// LS Electric XG5000 project: COMFactoryIO_Automated Warehouse10TL
// PLC LSPLC

PROGRAM NewProgram (task: 스캔 프로그램)

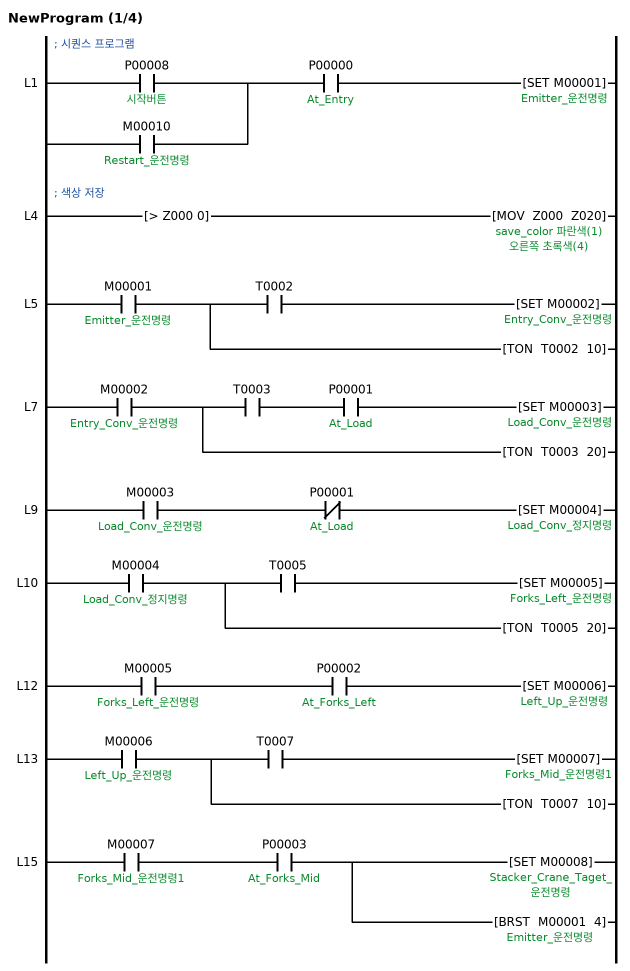
// 시퀀스 프로그램
; L1
LOAD      P00008	// 시작버튼
OR        M00010	// Restart_운전명령
AND       P00000	// At_Entry
SET       M00001	// Emitter_운전명령
// 색상 저장
; L4
LOAD>     Z000 0
MOV       Z000 Z020	// save_color 파란색(1) 오른쪽 초록색(4)
; L5
LOAD      M00001	// Emitter_운전명령
MPUSH
AND       T0002
SET       M00002	// Entry_Conv_운전명령
MPOP
TON       T0002 10
; L7
LOAD      M00002	// Entry_Conv_운전명령
MPUSH
AND       T0003
AND       P00001	// At_Load
SET       M00003	// Load_Conv_운전명령
MPOP
TON       T0003 20
; L9
LOAD      M00003	// Load_Conv_운전명령
AND NOT   P00001	// At_Load
SET       M00004	// Load_Conv_정지명령
; L10
LOAD      M00004	// Load_Conv_정지명령
MPUSH
AND       T0005
SET       M00005	// Forks_Left_운전명령
MPOP
TON       T0005 20
; L12
LOAD      M00005	// Forks_Left_운전명령
AND       P00002	// At_Forks_Left
SET       M00006	// Left_Up_운전명령
; L13
LOAD      M00006	// Left_Up_운전명령
MPUSH
AND       T0007
SET       M00007	// Forks_Mid_운전명령1
MPOP
TON       T0007 10
; L15
LOAD      M00007	// Forks_Mid_운전명령1
AND       P00003	// At_Forks_Mid
SET       M00008	// Stacker_Crane_Taget_운전명령
BRST      M00001 4	// Emitter_운전명령

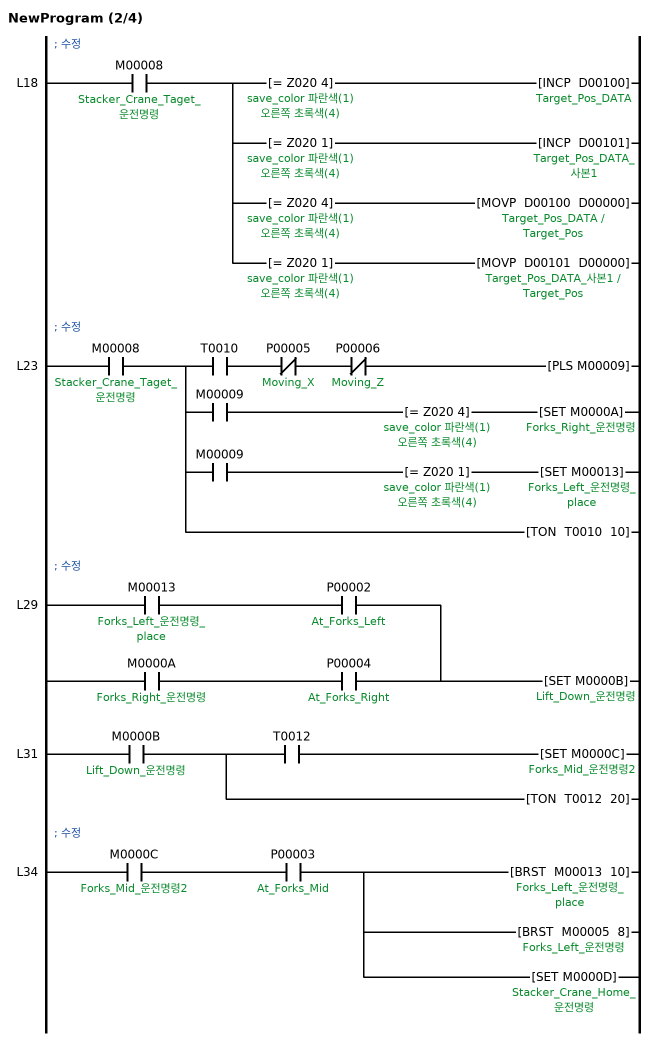
// 수정
; L18
LOAD      M00008	// Stacker_Crane_Taget_운전명령
MPUSH
AND=      Z020 4	// save_color 파란색(1) 오른쪽 초록색(4)
INCP      D00100	// Target_Pos_DATA
MLOAD
AND=      Z020 1	// save_color 파란색(1) 오른쪽 초록색(4)
INCP      D00101	// Target_Pos_DATA_사본1
MLOAD
AND=      Z020 4	// save_color 파란색(1) 오른쪽 초록색(4)
MOVP      D00100 D00000	// Target_Pos_DATA / Target_Pos
MPOP
AND=      Z020 1	// save_color 파란색(1) 오른쪽 초록색(4)
MOVP      D00101 D00000	// Target_Pos_DATA_사본1 / Target_Pos
// 수정
; L23
LOAD      M00008	// Stacker_Crane_Taget_운전명령
MPUSH
AND       T0010
AND NOT   P00005	// Moving_X
AND NOT   P00006	// Moving_Z
OUTP      M00009
MLOAD
AND       M00009
AND=      Z020 4	// save_color 파란색(1) 오른쪽 초록색(4)
SET       M0000A	// Forks_Right_운전명령
MLOAD
AND       M00009
AND=      Z020 1	// save_color 파란색(1) 오른쪽 초록색(4)
SET       M00013	// Forks_Left_운전명령_place
MPOP
TON       T0010 10
// 수정
; L29
LOAD      M00013	// Forks_Left_운전명령_place
AND       P00002	// At_Forks_Left
LOAD      M0000A	// Forks_Right_운전명령
AND       P00004	// At_Forks_Right
OR LOAD
SET       M0000B	// Lift_Down_운전명령
; L31
LOAD      M0000B	// Lift_Down_운전명령
MPUSH
AND       T0012
SET       M0000C	// Forks_Mid_운전명령2
MPOP
TON       T0012 20
// 수정
; L34
LOAD      M0000C	// Forks_Mid_운전명령2
AND       P00003	// At_Forks_Mid
BRST      M00013 10	// Forks_Left_운전명령_place
BRST      M00005 8	// Forks_Left_운전명령
SET       M0000D	// Stacker_Crane_Home_운전명령

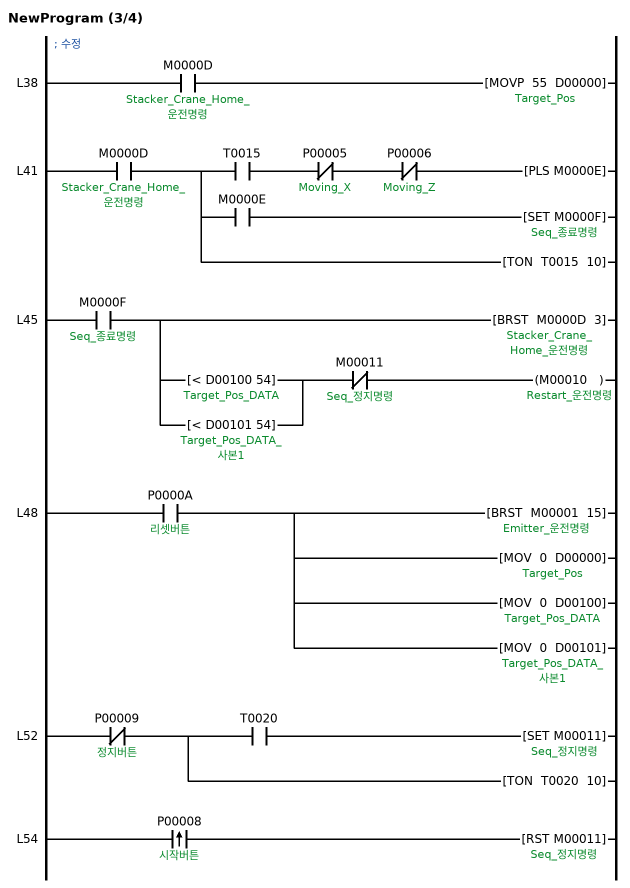
// 수정
; L38
LOAD      M0000D	// Stacker_Crane_Home_운전명령
MOVP      55 D00000	// Target_Pos
; L41
LOAD      M0000D	// Stacker_Crane_Home_운전명령
MPUSH
AND       T0015
AND NOT   P00005	// Moving_X
AND NOT   P00006	// Moving_Z
OUTP      M0000E
MLOAD
AND       M0000E
SET       M0000F	// Seq_종료명령
MPOP
TON       T0015 10
; L45
LOAD      M0000F	// Seq_종료명령
BRST      M0000D 3	// Stacker_Crane_Home_운전명령
LOAD<     D00100 54	// Target_Pos_DATA
OR<       D00101 54	// Target_Pos_DATA_사본1
AND LOAD
AND NOT   M00011	// Seq_정지명령
OUT       M00010	// Restart_운전명령
; L48
LOAD      P0000A	// 리셋버튼
BRST      M00001 15	// Emitter_운전명령
MOV       0 D00000	// Target_Pos
MOV       0 D00100	// Target_Pos_DATA
MOV       0 D00101	// Target_Pos_DATA_사본1
; L52
LOAD NOT  P00009	// 정지버튼
MPUSH
AND       T0020
SET       M00011	// Seq_정지명령
MPOP
TON       T0020 10
; L54
LOADP     P00008	// 시작버튼
RST       M00011	// Seq_정지명령

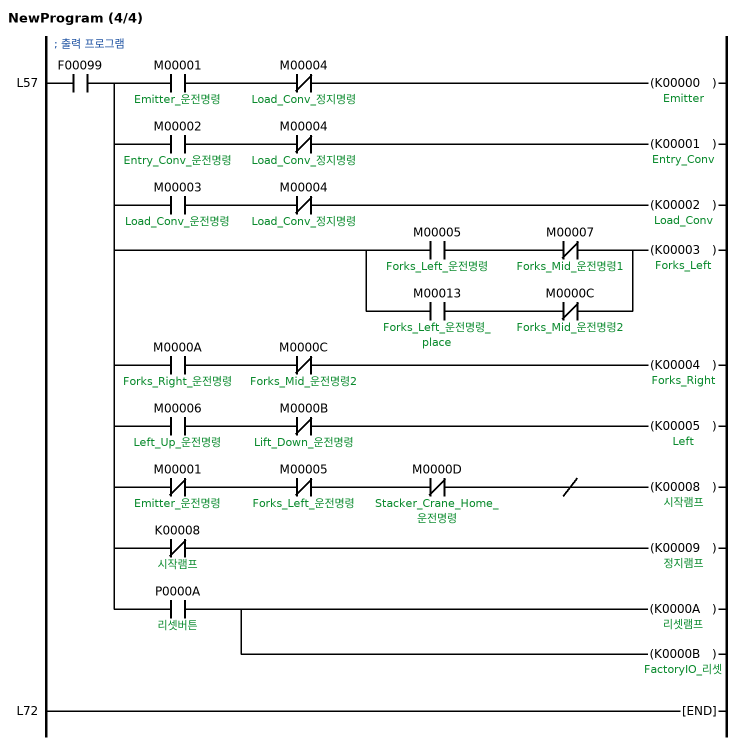
// 출력 프로그램
; L57
LOAD      F00099
MPUSH
AND       M00001	// Emitter_운전명령
AND NOT   M00004	// Load_Conv_정지명령
OUT       K00000	// Emitter
MLOAD
AND       M00002	// Entry_Conv_운전명령
AND NOT   M00004	// Load_Conv_정지명령
OUT       K00001	// Entry_Conv
MLOAD
AND       M00003	// Load_Conv_운전명령
AND NOT   M00004	// Load_Conv_정지명령
OUT       K00002	// Load_Conv
MLOAD
LOAD      M00005	// Forks_Left_운전명령
AND NOT   M00007	// Forks_Mid_운전명령1
LOAD      M00013	// Forks_Left_운전명령_place
AND NOT   M0000C	// Forks_Mid_운전명령2
OR LOAD
AND LOAD
OUT       K00003	// Forks_Left
MLOAD
AND       M0000A	// Forks_Right_운전명령
AND NOT   M0000C	// Forks_Mid_운전명령2
OUT       K00004	// Forks_Right
MLOAD
AND       M00006	// Left_Up_운전명령
AND NOT   M0000B	// Lift_Down_운전명령
OUT       K00005	// Left
MLOAD
AND NOT   M00001	// Emitter_운전명령
AND NOT   M00005	// Forks_Left_운전명령
AND NOT   M0000D	// Stacker_Crane_Home_운전명령
NOT
OUT       K00008	// 시작램프
MLOAD
AND NOT   K00008	// 시작램프
OUT       K00009	// 정지램프
MPOP
AND       P0000A	// 리셋버튼
OUT       K0000A	// 리셋램프
OUT       K0000B	// FactoryIO_리셋
; L72
END

VARIABLES AND COMMENTS (devices not used above)
D00001	WORD	Target_Pos_사본1
M00000	BIT	운전중